Fanuc KAREL source: kt00338.KL

-- PROVISIONAL review KL for V1013-1; original PC SHA256 a68ef51089ef39284fc3dd396f21fa100d07ebd0b966a9a0779fda2f797e2b26
-- Incomplete behavior may be omitted. Consult companion uncertainty JSON. Do not deploy.
PROGRAM KT00338
%NOLOCKGROUP
VAR
  S1 : STRING[80]
  S2 : STRING[80]
  OUT : BOOLEAN
BEGIN
  -- UNRESOLVED_PC offsets 5-14; opcodes 3F,75
  -- UNRESOLVED_PC offsets 19-28; opcodes 3F,75
  -- UNRESOLVED_PC offsets 33-42; opcodes 3F,75
  -- UNRESOLVED_PC offsets 47-56; opcodes 3F,75
  -- UNRESOLVED_PC offsets 61-80; opcodes 73,73,85,23
  -- UNRESOLVED_PC offsets 85-89; opcodes 7F
END KT00338
